{attribute 'qualified_only'}
VAR_GLOBAL
	
	// BistableSingleCoilRelay ToggleVirtualState
	// Manually toggle internal, virtual relay state when mismatch with real, physical	
	Shutter1OpenRelayToggle : BOOL := FALSE;
	Shutter1CloseRelayToggle : BOOL := FALSE;
	
	// Shutters
	Shutter1CmdEvent : stShutterCmdEvent;
	Shutter1Position : stShutterPosition;
    Shutter1State : eShutterStateType;
	ShutterUpSavedPos : stShutterPosition;
	ShutterDownSavedPos : stShutterPosition;
	
	// Schedulerr
	Shutter1EveningScheduleSet : BOOL := FALSE;
END_VAR

VAR_GLOBAL RETAIN
	
	// Schedulers
	ScheduleMonths   : ARRAY[1..12] OF BOOL := [1, 1, 1, 1, 1, 1, 1, 1, 1, 1, 1, 1];
	ScheduleWeekDays : ARRAY[1..7] OF BOOL := [1, 1, 1, 1, 1, 1, 1];
    ScheduleTimes    : ARRAY[1..6] OF TIME_OF_DAY := [
        TOD#17:10,
        TOD#17:15,
        TOD#17:20,
        TOD#17:25,
        TOD#00:00,
        TOD#00:00
    ];

	Shutter1EveningScheduleConfig : stSchedulerConfig := (Months := ScheduleMonths,
															WeekDays := ScheduleWeekDays,
															Times := ScheduleTimes);
END_VAR

(* stored: Version 1.1.0.1
   GVL gvlHA: Id {0181db7e-994c-475a-978f-c286ac6dc635} *)
